Staubli VAL3: cycle_Abort.pgx

program cycle_Abort()
begin
  // abort task
  rs:_nOmacStat=10
  taskKill("GoHome")
  taskKill("Monitor")
  taskKill("RotGoHome")
  taskKill("Monitor1")
  call ar:getCurMoveID(bGetMovId,"Abort")
  stopMove()
  resetMotion()

  // Stop task
  taskKill("Reset")
  taskKill("Start")
  taskKill("Stop")
  taskKill("End")
  taskKill("productCycle")
  taskKill("getForce")
  wait(isSettled())
  disablePower()
  wait(isPowered()==false)
    //2025.7.21 add 复位输出信号
  call plc:resetOutput()
  //OMAC进程:Stopped
  rs:_nOmacStat=9
  logMsg("当前处于生产停止状态 "+toString(".2",clock()))
  rs:_sRobotStatus="当前处于生产停止状态"
  delay(0)
end
